(* IEC 61131-3 sources: 89152_FlorisHendrix_AfstudeerProject/89152_FlorisHendrix_ExamenProject/Stations/MachineControl/MachineControl/Class/TCPCommunication (part 2) *)

      udAliveError := ParaVal$UDINT;

    //**************************************************************************
    TCPCom_ParaWR_AliveSignalTime: // - SET TIME FOR SENDING ALIVE SIGNAL -
    //**************************************************************************

      sParameter.udTimeAliveSignal := ParaVal$UDINT;

    //**************************************************************************
    TCPCOM_ParaWR_TaskPriority: // - SET TASK PRIORITY FOR THE TCP TASK -
    //**************************************************************************

      uiTaskPriority := ParaVal$UINT;

    // KruAle v1.16: Set timeout for sending Acknowledge and KeepAlive Messages
    //**************************************************************************
    TCPCOM_ParaWR_AckSendTimeout: // - SET TIMEOUT FOR ACK-MSG AND ALIVE-MSG -
    //**************************************************************************

      sParameter.udTimeOutAlive := ParaVal$UDINT;

    // KruAle v1.16: Set number of retries for sending Acknowledge and KeepAlive Messages
    //**************************************************************************
    TCPCOM_ParaWR_AckSendRetries: // - SET RETRIES FOR ACK-MSG AND ALIVE-MSG -
    //**************************************************************************

      // Max. Retries is 255
      if ParaVal > 0xFF then
        ParaVal := 0xFF;
      end_if;
      usRetriesAckTimeout := ParaVal$USINT;

    // KruAle v1.16: Set error-handling for sending Acknowledge and KeepAlive Messages
    //**************************************************************************
    TCPCOM_ParaWR_AckErrCloseConn: // - SET ERROR HANDLING FOR ACK-MSG -
    //**************************************************************************

      bAckErrorCloseConnection := ParaVal$BOOL;

    //**************************************************************************
    else // - INVALID PARAMETER NUMBER
    //**************************************************************************

      Retcode := -1001;

  end_case;

END_FUNCTION

FUNCTION GLOBAL TCPCommunication::ReadParameter
VAR_INPUT
  ParaNo 	  : DINT;
  pParaVal 	: ^DINT;
END_VAR
VAR_OUTPUT
  Retcode 	: DINT;
END_VAR

  Retcode := 0;

  if (pParaVal = NIL) then
    Retcode := -1002;
  end_if;

  case ParaNo of

    //**************************************************************************
    TCPCom_ParaRD_ComPort: // - READ COM PORT -
    //**************************************************************************

      pParaVal^$UDINT := ComPort;

    //20170410 DacPat v1.9 Added ReadParameter for the time interval between each transferrate calculation and each send alive signal
    //**************************************************************************
    TCPCom_ParaRD_MissingAliveError: // - READ ERROR THRESHOLD FOR ALIVE SIG -
    //**************************************************************************

      pParaVal^$UDINT := udAliveError;

    //**************************************************************************
    TCPCom_ParaRD_AliveSignalTime: // - READ TIME FOR SENDING ALIVE SIGNAL -
    //**************************************************************************

      pParaVal^$UDINT := sParameter.udTimeAliveSignal;

    //**************************************************************************
    TCPCom_ParaRD_TaskPriority: // - READ TASK PRIORITY FOR THE TCP TASK -
    //**************************************************************************

      pParaVal^$UINT := uiTaskPriority;

    // KruAle v1.15: Added ReadParameter to read the size of the send buffer
    //**************************************************************************
    TCPCom_ParaRD_TCPSendBuffersize: // - READ SIZE OF SEND BUFFER -
    //**************************************************************************

      pParaVal^$UDINT := udAllocSendBuffersize;

    // KruAle v1.16: Get timeout for sending Acknowledge and KeepAlive Messages
    //**************************************************************************
    TCPCOM_ParaRD_AckSendTimeout: // - READ TIMEOUT FOR ACK-MSG AND ALIVE-MSG -
    //**************************************************************************

      pParaVal^$UDINT := sParameter.udTimeOutAlive;

    // KruAle v1.16: Get number of retries for sending Acknowledge and KeepAlive Messages
    //**************************************************************************
    TCPCOM_ParaRD_AckSendRetries: // - READ RETRIES FOR ACK-MSG AND ALIVE-MSG -
    //**************************************************************************

      pParaVal^$USINT := usRetriesAckTimeout;

    // KruAle v1.16: Read error-handling for sending Acknowledge and KeepAlive Messages
    //**************************************************************************
    TCPCOM_ParaRD_AckErrCloseConn: // - READ ERROR HANDLING FOR ACK-MSG -
    //**************************************************************************

      pParaVal^$BOOL := bAckErrorCloseConnection;

    //**************************************************************************
    else // - INVALID PARAMETER NUMBER
    //**************************************************************************

      Retcode := -1001;

  end_case;

END_FUNCTION

FUNCTION TCPCommunication::ComStop
VAR_OUTPUT
  Retcode 	: DINT;
END_VAR

  Retcode := 0;

  sConfig.bComDeactivated := true;

  if (eComSteps > TCPCom_StartConnecting) then
    eComSteps := TCPCom_CloseConnection;
  else
    eComSteps := TCPCom_Deactivated;
  end_if;

END_FUNCTION

FUNCTION TCPCommunication::ComStart
VAR_OUTPUT
  Retcode 	: DINT;
END_VAR

  Retcode := 0;

  sConfig.bComDeactivated  := false;

END_FUNCTION

FUNCTION VIRTUAL GLOBAL TCPCommunication::DeactivateCom::Write
VAR_INPUT
  input (EAX) 	: DINT;
END_VAR
VAR_OUTPUT
  result (EAX) 	: DINT;
END_VAR
VAR
	dRet          : DINT;
END_VAR

  case DeactivateCom of

    //*****************************************************************************
    0: // - COMMUNICATION IS ACTIVATED
    //*****************************************************************************
      if (input = 1) then
        dRet := ComStop();
        if (dRet = 0) then
          DeactivateCom := input;
          result := DeactivateCom;
        else
          result := ACCESS_DENIED;
        end_if;
      else
        result := DeactivateCom;
      end_if;

    //*****************************************************************************
    1: // - COMMUNICATION IS DEACTIVATED
    //*****************************************************************************
      if (input = 0) then
        dRet := ComStart();
        if (dRet = 0) then
          DeactivateCom := input;
          result := DeactivateCom;
        else
          result := ACCESS_DENIED;
        end_if;
      else
        result := DeactivateCom;
      end_if;

  end_case;

END_FUNCTION

#define DESTPLC_WINPC_98    0x000001B // LARS, Standard PC, Win98/ME
#define DESTPLC_WINPC_NT    0x000001C // LARS, Standard PC, WinNT/Win2000/WinXP
#define DESTPLC_WINIPC_98   0x000001D // LARS, IPC, Win98/ME
#define DESTPLC_WINIPC_NT   0x000001E // LARS, IPC, WinNT/Win2000/WinXP

FUNCTION TCPCommunication::IsLars
	VAR_OUTPUT
		retcode 	: DINT;
	END_VAR

  retcode := FALSE;
  case _WHOAMI of
    DESTPLC_WINPC_98,
    DESTPLC_WINPC_NT,
    DESTPLC_WINIPC_98,
    DESTPLC_WINIPC_NT : retcode := TRUE;
  end_case;

END_FUNCTION

FUNCTION TCPCommunication::DelayComTask
	VAR_INPUT
		udDelay 	: UDINT;
	END_VAR

  if IsSalamanderOS = TRUE then
    OSSD_DELAY(pCIL_DEBUG, udDelay*1000); // Microseconds!
  else
    coMultiTask.TASKDELAY(udDelay);
  end_if;

END_FUNCTION
